Fanuc KAREL source: kf00114.KL

-- PROVISIONAL review KL for V1013-1; original PC SHA256 2328c929dee85e31db0c47b2b48124644181a770c294fdbc5b862775fa09b0ee
-- Incomplete behavior may be omitted. Consult companion uncertainty JSON. Do not deploy.
PROGRAM KF00114
%NOLOCKGROUP
BEGIN
  -- UNRESOLVED_PC offsets 0-1; opcodes 7B
  -- UNRESOLVED_PC offsets 6-20; opcodes 2D,9D,52,23
  -- UNRESOLVED_PC offsets 25-29; opcodes 7F
  -- UNRESOLVED_PC offsets 34-44; opcodes 27,22,AA
  -- UNRESOLVED_PC offsets 49-53; opcodes 7F
END KF00114
